Fanuc KAREL source: kb00181.KL

-- PROVISIONAL review KL for V940-1; original PC SHA256 a2b01030a8d05f7ea5b217d06e1edc3516ccff5ae40bff3bdfb22f8047c27942
-- Incomplete behavior may be omitted. Consult companion uncertainty JSON. Do not deploy.
PROGRAM KB00181
%NOLOCKGROUP
BEGIN
  -- V9_ZERO_TABLE_METADATA_HINT layout=0002_ascii; no indexed target words; source/name/runtime held
  -- UNRESOLVED_PC offsets 5-12; opcodes 9D,23
  -- UNRESOLVED_PC offsets 17-27; opcodes 27,22,31
  -- UNRESOLVED_PC offsets 32-36; opcodes 7F
END KB00181
